// TIA Portal V21 export
// export: Created 2000-01-01T00:00:00.0000000Z, ExportSetting None
TYPE "UDT_HMI_DualEStop"
   STRUCT
      bHmiResetCmd { ExternalWritable := 'False'} : Bool;   // HMI安全复位请求（须配合现场双通道正常）
      tDiscrepancyTime { ExternalWritable := 'False'} : Time;   // 双通道不同步最大允许差异时间（默认 T#200ms）
      bSafeToRun { ExternalWritable := 'False'} : Bool;   // 状态反馈：安全回路已闭合允许运行
      bCh1State { ExternalWritable := 'False'} : Bool;   // 状态反馈：急停通道1状态
      bCh2State { ExternalWritable := 'False'} : Bool;   // 状态反馈：急停通道2状态
      bDiscrepancyFault { ExternalWritable := 'False'} : Bool;   // 状态反馈：双通道不一致触点粘连故障
      bWaitReset { ExternalWritable := 'False'} : Bool;   // 状态反馈：等待人工复位脉冲
      wStatus { ExternalWritable := 'False'} : Word;   // 状态码：16#0000安全闭合, 16#7001等待复位, 16#8401急停按下, 16#8402安全门打开, 16#8403双通道不同步故障
   END_STRUCT;
END_TYPE
